// TIA Portal V21 export
// export: Created 2026-11-10T19:12:26.7955029Z, ExportSetting WithDefaults, DisplayName Totally Integrated Automation Portal, DisplayVersion V21 Update 3, DisplayName STEP 7 Professional, DisplayVersion V21 Update 3, DisplayName STEP 7 Safety, DisplayVersion V21, DisplayName Tech WebApplication, DisplayVersion V21, DisplayName WinCC Basic/Comfort/Advanced, DisplayVersion V21 Update 3, DisplayName WinCC Unified, DisplayVersion V21 Update 3
DATA_BLOCK "DBsTCONT_S"   // DB34
// stored: AutoNumber true, DBAccessibleFromOPCUA true, DBAccessibleFromWebserver true, InstanceOfName TCONT_S, OfSystemLibElement TCONT_S, OfSystemLibVersion 1.1
TCONT_S   // technology object, version 1.1
   // VAR_INPUT
   //    CYCLE : Real;
   //    SP_INT : Real;
   //    PV_IN : Real;
   //    PV_PER : Int;
   //    DISV : Real;
   //    LMNR_HS : Bool;
   //    LMNR_LS : Bool;
   //    LMNS_ON : Bool;
   //    LMNUP : Bool;
   //    LMNDN : Bool;
   // END_VAR
   // VAR_OUTPUT
   //    QLMNUP : Bool;
   //    QLMNDN : Bool;
   //    PV : Real;
   //    ER : Real;
   // END_VAR
   // VAR_IN_OUT
   //    COM_RST : Bool;
   // END_VAR
   // VAR RETAIN
   //    PV_FAC : Real;
   //    PV_OFFS : Real;
   //    DEADB_W : Real;
   //    PFAC_SP : Real;
   //    GAIN : Real;
   //    TI : Real;
   //    MTR_TM : Real;
   //    PULSE_TM : Real;
   //    BREAK_TM : Real;
   //    PER_MODE : Int;
   //    PVPER_ON : Bool;
   //    sFbPVal : Real;
   //    sThrOn : Real;
   //    siImpAus : Int;
   //    stImpDauer : Real;
   //    stPausDauer : Real;
   //    srSpOld : Real;
   //    srDiffSp : Real;
   // END_VAR
BEGIN
END_DATA_BLOCK
